TYPE ST_VC_ReportModuleStateArgs :
STRUCT
    State   : UINT;     // PackML state from VisionCore
    AlarmId : DINT;
END_STRUCT
END_TYPE

(* stored: Version 1.1.0.1, ProductVersion 3.1.4026.21
   DUT ST_VC_ReportModuleStateArgs: Id {a79ef6cb-a06e-4d2a-a3a7-3fd26c1d581f} *)
